{attribute 'no_assign'}
FUNCTION_BLOCK FB_LN_WTURBINE_LD0_WALM1 EXTENDS FB_AcsiCommonLogicalNodeClass
VAR_INPUT
	Beh: FB_DO_WTURBINE_LD0_WALM1_Beh := (sClass:='ENS', bLinkResult:=THIS^.AddDataToContainer(ipData:=Beh));
END_VAR
VAR
END_VAR

END_FUNCTION_BLOCK

(* stored: Version 1.1.0.1
   POU FB_LN_WTURBINE_LD0_WALM1: Id {21b07012-2fad-47e4-a5d5-b3a26da7c962}, SpecialFunc None *)
